(*
SPDX-FileCopyrightText: c 2026 Oleksandr Tiutyk <trofimich@gmail.com>
SPDX-License-Identifier: MIT
License: https://opensource.org/license/mit
*)

(*!
<summary>Checks ANY lookup after growth and head removal.</summary>
<description>
Owns a dynamic queue and copied payloads at a stable address. Run from one task.
Teardown clears surviving entries and releases dynamic capacity.
</description>
*)

{attribute 'no_assign'}
{attribute 'no_explicit_call' := 'do not call this function block directly'}
FUNCTION_BLOCK DynamicQueueContainsTest EXTENDS TOF_Testing.SingleCycleTest
VAR_STAT
	{attribute 'hide'}
	_ClassName : STRING := __POUNAME();
END_VAR
VAR
	_Queue : TOF_Collections.Queue<0>(valueValidator := 0);
END_VAR

(*!
<summary>Checks ANY lookup after growth and head removal.</summary>
*)
METHOD PROTECTED ExecuteTest
VAR
	values : ARRAY [1..4] OF INT := [11, 22, 33, 44];
END_VAR
_Queue.DefaultDynamicAllocationElementCount := BYTE#2;

_Queue
	.EnqueueCopy(value := values[1])
	.EnqueueCopy(value := values[2])
	.EnqueueCopy(value := values[3]);

Assert.ThatBool(
	actual := _Queue.Contains(value := values[1]),
	message := "Lookup must find the original head after growth"
).IsTrue();

Assert.ThatBool(
	actual := _Queue.Contains(value := values[3]),
	message := "Lookup must find the entry appended during growth"
).IsTrue();

Assert.ThatBool(
	actual := _Queue.Contains(value := values[4]),
	message := "Lookup must reject an absent value"
).IsFalse();

_Queue.RemoveFirst();

Assert.ThatBool(
	actual := _Queue.Contains(value := values[1]),
	message := "Lookup must ignore the removed head"
).IsFalse();

Assert.ThatDInt(
	actual := _Queue.Length,
	message := "Lookup must preserve the two live entries"
).ToBe(expected := DINT#2);

Assert.ThatInt(
	actual := _Queue.Peek().AsInt(),
	message := "Lookup must preserve the current head"
).ToBe(expected := values[2]);
END_METHOD

(*!
<summary>Clears the fixture before the runner publishes the result.</summary>
<description>
Also runs after an unexpected exception interrupts the case.
</description>
*)
METHOD PROTECTED AfterTest
_Queue.Clear();
END_METHOD

//! <summary>Borrows the concrete class name. Callers must not modify it.</summary>
{attribute 'monitoring' := 'call'}
PROPERTY ClassName : REFERENCE TO STRING
GET
ClassName REF= _ClassName;
END_GET
END_PROPERTY

//! <summary>Borrows the compiler-initialized namespace name. Callers must not modify it.</summary>
{attribute 'monitoring' := 'call'}
PROPERTY NamespaceName : REFERENCE TO STRING
GET
NamespaceName REF= CurrentNamespace.Name;
END_GET
END_PROPERTY

//! <summary>Reports the concrete instance size in bytes.</summary>
{attribute 'monitoring' := 'call'}
PROPERTY SelfSize : ULINT
GET
SelfSize := XSIZEOF(THIS^);
END_GET
END_PROPERTY

END_FUNCTION_BLOCK

(* stored: Version 1.1.0.1
   POU DynamicQueueContainsTest: Id {94bb8e6f-b8f9-4f1a-9f04-fb780f2c6c2f}, SpecialFunc None
   Method ExecuteTest: Id {6abcb50c-c270-4be6-9fdc-38cecb20f192}
   Method AfterTest: Id {fd80e976-1bbf-4965-898d-ce8f0f102452}
   Property ClassName: Id {12b793f0-1e39-480d-a6cb-2792b4ed722c}
   Get Get: Id {916ea62f-9958-496a-bc2f-45e5e60f2863}
   Property NamespaceName: Id {41172de2-f9c3-4d48-bb70-c69023c8c886}
   Get Get: Id {da090ed5-45ef-445b-bf1d-a68ca2ca3560}
   Property SelfSize: Id {b0b2ced1-f1c5-41a5-8eed-22deb2e8f905}
   Get Get: Id {ce118f90-d79c-48ea-9623-108ac7594369} *)
